(* IEC 61131-3 sources: codesys-to-s7/tests/corpus/C2S7-TYPE-WSTRING/pos, 1 file *)

(* ---- input.st ---- *)
FUNCTION_BLOCK FB_Case
VAR
    ws : WSTRING;
END_VAR
ws := "a";
END_FUNCTION_BLOCK
